(* IEC 61131-3 sources: PortalRobot/Portal_robot/Device/application/ST/ST_MAGAZINE/ST_DETAIL, 2 files *)

(* ---- E_DETAIL_TYPE.st ---- *)
{attribute 'qualified_only'}
{attribute 'strict'}
TYPE E_DETAIL_TYPE :
(
	NONE,
	BLANK,
	DETAIL
);
END_TYPE

(* ---- ST_DETAIL.st ---- *)
TYPE ST_DETAIL :
STRUCT
	eDetailType : E_DETAIL_TYPE; // Тип содержимого слота
	xInPosition : BOOL; // Признак наличия объекта в слоте
	uiProductType : UINT; // Тип продукции перемещается между зонами вместе со слотом
END_STRUCT
END_TYPE
